// TIA Portal V17 export
// export: Created 2026-11-17T10:42:02.9478916Z, ExportSetting WithDefaults, DisplayName Totally Integrated Automation Portal, DisplayVersion V17, DisplayName TIA Portal Openness, DisplayVersion V17, DisplayName TIA Portal Version Control Interface, DisplayVersion V17, DisplayName STEP 7 Professional, DisplayVersion V17, DisplayName STEP 7 Safety, DisplayVersion V17, DisplayName WinCC Advanced, DisplayVersion V17
ORGANIZATION_BLOCK "Main"   // OB1, LAD, ProgramCycle
{ S7_Optimized_Access := 'TRUE' }
VERSION : 0.1
// stored: AutoNumber true, IsIECCheckEnabled false, SetENOAutomatically false
   VAR_INPUT
      Initial_Call : Bool;   // Initial call of this OB
      Remanence : Bool;   // =True, if remanent data are available
   END_VAR
BEGIN

REGION Network 1: 启停自锁
   // 启动后保持运行，停止优先。
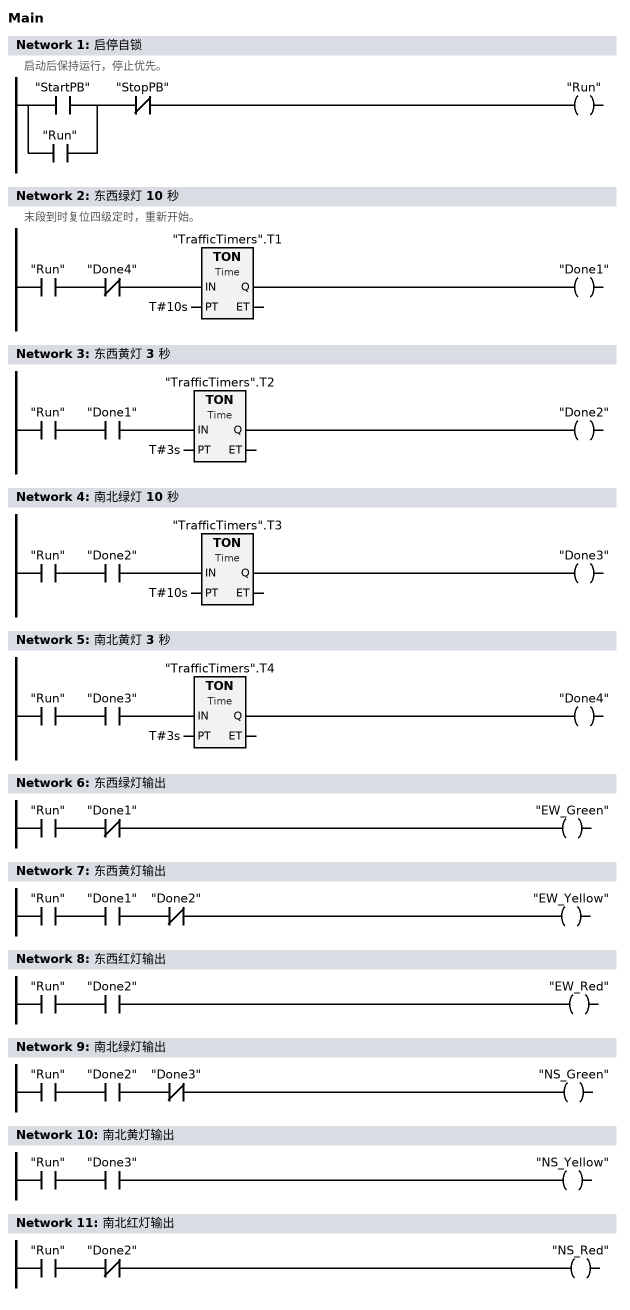
   RUNG wire#powerrail
      Contact( "StartPB" )
      wire#w1
      I_Contact( "StopPB" )
      Coil( "Run" )
   END_RUNG
   RUNG wire#powerrail
      Contact( "Run" )
   END_RUNG wire#w1
   // the same network as SCL:
   "Run" := ("StartPB" OR "Run") AND NOT "StopPB";
END_REGION

REGION Network 2: 东西绿灯 10 秒
   // 末段到时复位四级定时，重新开始。
   RUNG wire#powerrail
      Contact( "Run" )
      I_Contact( "Done4" )
      { S7_Templates := "time_type := Time" } "TrafficTimers".T1.TON(pt := T#10s, et =>)
      Coil( "Done1" )
   END_RUNG
   // the same network as SCL:
   "TrafficTimers".T1.TON(IN := "Run" AND NOT "Done4", PT := T#10s);
   "Done1" := "TrafficTimers".T1.Q;
END_REGION

REGION Network 3: 东西黄灯 3 秒
   RUNG wire#powerrail
      Contact( "Run" )
      Contact( "Done1" )
      { S7_Templates := "time_type := Time" } "TrafficTimers".T2.TON(pt := T#3s, et =>)
      Coil( "Done2" )
   END_RUNG
   // the same network as SCL:
   "TrafficTimers".T2.TON(IN := "Run" AND "Done1", PT := T#3s);
   "Done2" := "TrafficTimers".T2.Q;
END_REGION

REGION Network 4: 南北绿灯 10 秒
   RUNG wire#powerrail
      Contact( "Run" )
      Contact( "Done2" )
      { S7_Templates := "time_type := Time" } "TrafficTimers".T3.TON(pt := T#10s, et =>)
      Coil( "Done3" )
   END_RUNG
   // the same network as SCL:
   "TrafficTimers".T3.TON(IN := "Run" AND "Done2", PT := T#10s);
   "Done3" := "TrafficTimers".T3.Q;
END_REGION

REGION Network 5: 南北黄灯 3 秒
   RUNG wire#powerrail
      Contact( "Run" )
      Contact( "Done3" )
      { S7_Templates := "time_type := Time" } "TrafficTimers".T4.TON(pt := T#3s, et =>)
      Coil( "Done4" )
   END_RUNG
   // the same network as SCL:
   "TrafficTimers".T4.TON(IN := "Run" AND "Done3", PT := T#3s);
   "Done4" := "TrafficTimers".T4.Q;
END_REGION

REGION Network 6: 东西绿灯输出
   RUNG wire#powerrail
      Contact( "Run" )
      I_Contact( "Done1" )
      Coil( "EW_Green" )
   END_RUNG
   // the same network as SCL:
   "EW_Green" := "Run" AND NOT "Done1";
END_REGION

REGION Network 7: 东西黄灯输出
   RUNG wire#powerrail
      Contact( "Run" )
      Contact( "Done1" )
      I_Contact( "Done2" )
      Coil( "EW_Yellow" )
   END_RUNG
   // the same network as SCL:
   "EW_Yellow" := "Run" AND "Done1" AND NOT "Done2";
END_REGION

REGION Network 8: 东西红灯输出
   RUNG wire#powerrail
      Contact( "Run" )
      Contact( "Done2" )
      Coil( "EW_Red" )
   END_RUNG
   // the same network as SCL:
   "EW_Red" := "Run" AND "Done2";
END_REGION

REGION Network 9: 南北绿灯输出
   RUNG wire#powerrail
      Contact( "Run" )
      Contact( "Done2" )
      I_Contact( "Done3" )
      Coil( "NS_Green" )
   END_RUNG
   // the same network as SCL:
   "NS_Green" := "Run" AND "Done2" AND NOT "Done3";
END_REGION

REGION Network 10: 南北黄灯输出
   RUNG wire#powerrail
      Contact( "Run" )
      Contact( "Done3" )
      Coil( "NS_Yellow" )
   END_RUNG
   // the same network as SCL:
   "NS_Yellow" := "Run" AND "Done3";
END_REGION

REGION Network 11: 南北红灯输出
   RUNG wire#powerrail
      Contact( "Run" )
      I_Contact( "Done2" )
      Coil( "NS_Red" )
   END_RUNG
   // the same network as SCL:
   "NS_Red" := "Run" AND NOT "Done2";
END_REGION
END_ORGANIZATION_BLOCK
